(* IEC 61131-3 sources: codesys-framework/txt/application/ToDo/Hardware/IO/Camera/FB_Camera/Private, 8 files *)

(* ---- Monitor.method.st ---- *)
METHOD PRIVATE Monitor
VAR_INPUT
END_VAR
VAR_INST
	uiConnectionAttempts	: UINT;
	uiMaxConnectionAttempts	: UINT;
END_VAR

// --- BEGIN IMPLEMENTATION ---

uiMaxConnectionAttempts	:= 5;

CASE _iStateMonitor OF

	0 :	//Startup
		IF NOT _xError THEN
 		   _iStateMonitor := _iStateMonitor + 10;
		END_IF

	10 :  //Init timer
		uiConnectionAttempts	:= uiConnectionAttempts + 1;
		_tonMonitor.IN := FALSE;
		//Init connection
		_clientState.xEnable := FALSE;

		//Timer inactive and no active connection
		IF NOT _tonMonitor.Q AND NOT _clientState.xActive THEN
			IF _clientRead.xActive AND _clientWrite.xActive THEN
		   	   _iStateMonitor := _iStateMonitor + 10;
			END_IF
		END_IF

	20: //Make connection
		_clientState.xEnable := TRUE;

		//Active connection
		IF _clientState.xActive AND NOT _clientState.xError THEN
		   _iStateMonitor := _iStateMonitor + 10;
		END_IF
		//Error
		IF _clientState.xError THEN
		   _iStateMonitor := 1000;
		END_IF

	30: //Recheck
		_tonMonitor.IN := TRUE;
		//Init connection
		_clientState.xEnable := FALSE;
		//Connected
		_xConnected := TRUE;

		uiConnectionAttempts := 0;

		//error
		IF _tonMonitor.Q THEN
			_iStateMonitor := 0;
		END_IF

  1000: //Error
		_xError := _clientState.xError;
		_iErrorId := 0;
		_sError := CONCAT(_scSysPar.adress.sAddr,': CAMERA NO CONNECTION');
		_iStateMonitor := 1100;

  1100: //Init connected -> wait for reset
  		IF	uiConnectionAttempts < uiMaxConnectionAttempts
		THEN
			_xError := FALSE;
			_iStateMonitor := 0;
		END_IF
		_xConnected := FALSE;

END_CASE

(* ---- ProcessConnect.method.st ---- *)
METHOD PRIVATE ProcessConnect
VAR_INPUT
END_VAR

// --- BEGIN IMPLEMENTATION ---

_xBusy := TRUE;

CASE _iStateConnect OF

	0:  //Startup
		IF NOT _xError THEN
		   _iStateConnect := _iStateConnect + 10;
		END_IF

	10: //connect
		IF ConnectMethod() THEN
		   _iStateConnect := 50;
		END_IF

	50 :
		_iStateConnect := 0;
		_xDone := TRUE;
		_xBusy := FALSE;
		_eState := E_CameraStates.Standby;

END_CASE

(* ---- ProcessDisconnect.method.st ---- *)
METHOD PRIVATE ProcessDisconnect
VAR_INPUT
END_VAR

// --- BEGIN IMPLEMENTATION ---

_xBusy := TRUE;

CASE _iStateDisconnect OF

	0:  //Startup
		IF NOT _xError THEN
		   _iStateDisconnect := _iStateDisconnect + 10;
		END_IF

	10: //Init connection
		_clientRead.xEnable := FALSE;
		_clientWrite.xEnable := FALSE;

		//No active connections
		IF NOT _clientRead.xActive AND NOT _clientWrite.xActive THEN
		   _iStateDisconnect := _iStateDisconnect + 10;
		END_IF

	20 :
		_iStateDisconnect := 0;
		_xDone := TRUE;
		_xBusy := FALSE;
		_eState := E_CameraStates.Standby;

END_CASE

(* ---- ProcessFBs.method.st ---- *)
METHOD PRIVATE ProcessFBs
VAR_INPUT
END_VAR

// --- BEGIN IMPLEMENTATION ---

_clientRead(ipAddr := _scSysPar.adress,uiPort := _scSysPar.readPort,udiTimeOut := _scSysPar.conTimeout);
_clientWrite(ipAddr := _scSysPar.adress,uiPort := _scSysPar.writePort,udiTimeOut := _scSysPar.conTimeout);
_clientState(ipAddr := _scSysPar.adress,uiPort := _scSysPar.writePort,udiTimeOut := _scSysPar.conTimeout);

_read(
	xEnable:= _clientRead.xActive,
	xDone=> ,
	xBusy=> ,
	xError=> ,
	hConnection:= _clientRead.hConnection,
	szSize:= SIZEOF(_sResult),
	pData:= ADR(_sResult),
	eError=> ,
	xReady=> ,
	szCount=>
);

_write(
	xExecute:= ,
	udiTimeOut:= ,
	xDone=> ,
	xBusy=> ,
	xError=> ,
	hConnection:= _clientWrite.hConnection,
	szSize:= ,
	pData:= ,
	eError=>
);

_writeFeedBack(
	xEnable:= _clientWrite.xActive,
	xDone=> ,
	xBusy=> ,
	xError=> ,
	hConnection:= _clientWrite.hConnection,
	szSize:= SIZEOF(_sFeedBack),
	pData:= ADR(_sFeedBack),
	eError=> ,
	xReady=> ,
	szCount=>
);

_tonMonitor(PT := _scSysPar.monitorTime);
_tonPicture(PT := _scSysPar.readTimeout);
_tonSelectJob(PT := _scSysPar.jobTimeout);

(* ---- ProcessSelectJob.method.st ---- *)
METHOD PRIVATE ProcessSelectJob
VAR_INPUT
END_VAR
VAR
	result : STRING;
END_VAR

// --- BEGIN IMPLEMENTATION ---

_xBusy := TRUE;

CASE _iStateSetJob OF

	0 :
		_sJob := 'CJP00';
		_sJob := CONCAT('CJP00', UINT_TO_STRING(_id));
		_write.szSize := SIZEOF(_sJob);
		_write.pData := ADR(_sJob);
		_write.xExecute := TRUE;
		_tonSelectJob.IN := FALSE;

		_iStateSetJob := _iStateSetJob + 10;

	10 :
		_tonSelectJob.IN := TRUE;
		result := CONCAT('CJPPT00', UINT_TO_STRING(_id));

		IF _sFeedBack = result THEN
			_sFeedBack := '';
			_write.xExecute := FALSE;

			_xDone := TRUE;
			_eState := E_CameraStates.Standby;
			_iStateSetJob := 0;
		END_IF

		IF _tonSelectJob.Q THEN
			_iStateSetJob := 100;
		END_IF

	100 :
		_write.xExecute := FALSE;
		_iStateSetJob := _iStateSetJob + 10;

	110 :
		_iStateSetJob := 0;

END_CASE

(* ---- ProcessState.method.st ---- *)
METHOD PRIVATE ProcessState
VAR_INPUT
END_VAR

// --- BEGIN IMPLEMENTATION ---

CASE _eState OF

	E_CameraStates.None				: ;
	E_CameraStates.Invalid 			: _eState := E_CameraStates.Initialize;
	E_CameraStates.Initialize 		: Initialize();
	E_CameraStates.Connect 			: ProcessConnect();
	E_CameraStates.Disconnect 		: ProcessDisconnect();
	E_CameraStates.Standby 			: _xDone := FALSE; _xBusy := FALSE;
	E_CameraStates.SelectJob 		: ProcessSelectJob();
	E_CameraStates.TakePicture 		: ProcessTakePictureTRX();
	E_CameraStates.Reset 			: ProcessDisconnect();

END_CASE

(* ---- ProcessTakePicture.method.st ---- *)
METHOD PRIVATE ProcessTakePicture
VAR_INPUT
END_VAR
VAR
	result 	: STRING;
END_VAR

// --- BEGIN IMPLEMENTATION ---

_xBusy := TRUE;

CASE _iStateTakePicture OF

	0 :
		_sResult := '';
		_sPicture := 'ASH11';
		_write.szSize := SIZEOF(_sPicture);
		_write.pData := ADR(_sPicture);
		_write.xExecute := TRUE;

		_iStateTakePicture := _iStateTakePicture + 10;

	10 :
		IF Mid(STR := _sFeedBack, LEN := 4, POS := 1) = 'ASHP' THEN
			_sFeedBack := '';
			_write.xExecute := FALSE;
			_iStateTakePicture := _iStateTakePicture + 10;
		END_IF

	20 :
		//_tonPicture.IN := TRUE;

		//IF _tonPicture.Q THEN
			_tonPicture.IN := FALSE;
			_iStateTakePicture := _iStateTakePicture + 10;
		//END_IF

	30 :
		_sPicture := 'TRG';
		_write.szSize := SIZEOF(_sPicture);
		_write.pData := ADR(_sPicture);
		_write.xExecute := TRUE;

		_iStateTakePicture := _iStateTakePicture + 10;

	40 :
		IF _sFeedBack = 'TRGP' THEN
			_sFeedBack := '';
			_write.xExecute := FALSE;
			_iStateTakePicture := _iStateTakePicture + 10;
		ELSIF _sFeedBack = 'TRGF' THEN
			_sFeedBack := '';
			_write.xExecute := FALSE;
			_iStateTakePicture := 20;
		END_IF

	50 :
		_tonPicture.IN := TRUE;

		IF _tonPicture.Q and _sResult <> '' THEN
			_tonPicture.IN := FALSE;
			_iStateTakePicture := _iStateTakePicture + 10;
		END_IF

	60 :
		_iStateTakePicture := 0;
		_xDone := TRUE;
		_eState := E_CameraStates.Standby;

END_CASE

(* ---- ProcessTakePictureTRX.method.st ---- *)
METHOD PRIVATE ProcessTakePictureTRX
VAR_INPUT
END_VAR
VAR
	result 	: STRING;
END_VAR

// --- BEGIN IMPLEMENTATION ---

_xBusy := TRUE;

CASE _iStateTakePicture OF

	0 :
		_sResult := '';
		_sPicture := 'ASH11';
		_write.szSize := SIZEOF(_sPicture);
		_write.pData := ADR(_sPicture);
		_write.xExecute := TRUE;

		_iStateTakePicture := _iStateTakePicture + 10;

	10 :
		IF MID(STR := _sFeedBack, LEN := 4, POS := 1) = 'ASHP' THEN
			_sFeedBack := '';
			_write.xExecute := FALSE;
			_iStateTakePicture := _iStateTakePicture + 10;
		END_IF

	20 :
		//_tonPicture.IN := TRUE;

		//IF _tonPicture.Q THEN
			_tonPicture.IN := FALSE;
			_iStateTakePicture := _iStateTakePicture + 10;
		//END_IF

	30 :
		_sPicture := _sPictureId; //MID(STR := _sPictureId, LEN := 5, POS := 1);
		_write.szSize := SIZEOF(_sPicture);
		_write.pData := ADR(_sPicture);
		_write.xExecute := TRUE;

		_iStateTakePicture := _iStateTakePicture + 10;

	40 :
		IF MID(STR := _sFeedBack, LEN := 4, POS := 1) = 'TRXP' THEN
			_sFeedBack := '';
			_write.xExecute := FALSE;
			_iStateTakePicture := _iStateTakePicture + 10;
		ELSIF MID(STR := _sFeedBack, LEN := 4, POS := 1) = 'TRXF' THEN
			_sFeedBack := '';
			_write.xExecute := FALSE;
			_iStateTakePicture := 20;
		END_IF

	50 :
		_tonPicture.IN := TRUE;

		IF _tonPicture.Q and _sResult <> '' THEN
			_tonPicture.IN := FALSE;
			_iStateTakePicture := _iStateTakePicture + 10;
		END_IF

	60 :
		_iStateTakePicture := 0;
		_xDone := TRUE;
		_eState := E_CameraStates.Standby;

END_CASE
